(* IEC 61131-3 sources: stc/examples, 2 files *)

(* ---- inter.st ---- *)
(* Copyright (C) 2021-2026 Manuele Conti
   SPDX-License-Identifier: GPL-2.0-or-later
   Summary: Demonstrates function declarations, branching, typed values, and loops. *)

FUNCTION inter : INT
VAR_INPUT
    a_1: SINT;
    b_1: INT;
    test: BOOL;
END_VAR
VAR
    ff: INT;
END_VAR
    test := TRUE;
    IF a_1 = b_1 THEN
        a_1 := 70;
    ELSIF b_1 = 1 THEN
        b_1 := INT#10;
    END_IF;
    inter := a_1 + b_1;
    FOR ff := 1 TO 10 DO
	a_1 := a_1 + ff;
    END_FOR;
END_FUNCTION

(* ---- employee_oop.st ---- *)
(* Employee polymorphism inspired by:
   https://stefanhenneken.net/2020/12/13/iec-61131-3-abstract-fb-vs-interface/

   STC models the example with IEC Edition 3 CLASS declarations. Properties,
   REFERENCE TO and TwinCAT abstract FUNCTION_BLOCK extensions are deliberately
   replaced by fields, interfaces and methods supported by the compiler. *)

INTERFACE IEmployee
METHOD GetMonthlySalary : LREAL
END_METHOD
END_INTERFACE

CLASS ABSTRACT EmployeeBase IMPLEMENTS IEmployee
VAR
    EmployeeNumber : UINT;
END_VAR

METHOD PUBLIC ABSTRACT GetMonthlySalary : LREAL
END_METHOD

METHOD PUBLIC GetEmployeeNumber : UINT
    GetEmployeeNumber := EmployeeNumber;
END_METHOD
END_CLASS

CLASS FullTimeEmployee EXTENDS EmployeeBase
VAR
    AnnualSalary : LREAL;
END_VAR

METHOD PUBLIC OVERRIDE GetMonthlySalary : LREAL
    GetMonthlySalary := AnnualSalary / 12.0;
END_METHOD
END_CLASS

CLASS ContractEmployee EXTENDS EmployeeBase
VAR
    HourlyPay : LREAL;
    MonthlyHours : LREAL;
END_VAR

METHOD PUBLIC OVERRIDE GetMonthlySalary : LREAL
    GetMonthlySalary := HourlyPay * MonthlyHours;
END_METHOD
END_CLASS

PROGRAM EmployeeDemo
VAR
    FullTime : FullTimeEmployee;
    Contract : ContractEmployee;
    Employee : IEmployee;
    Salary : LREAL;
END_VAR
    FullTime.AnnualSalary := 120000.0;
    Contract.HourlyPay := 80.0;
    Contract.MonthlyHours := 160.0;

    Employee := FullTime;
    Salary := Employee.GetMonthlySalary();

    Employee := Contract;
    Salary := Employee.GetMonthlySalary();
END_PROGRAM
